(****************************************************************************************************<br>
© Syntegon Group.<br>
All rights reserved, also regarding any disposal, exploitation, reproduction, editing, distribution,<br>
as well as in the event of applications for industrial property rights.<br>
*****************************************************************************************************<br>
DESCRIPTION:<br>
Runtime-readable version of the Syn_Config library.<br>
*****************************************************************************************************<br>
VERSION         ¦ DATE       ¦ NAME      ¦ CHANGE<br>
Syn_Config 1.0.0 ¦ 2026-11-10 ¦ J.Willner ¦ Parameter sets of conveyors and Deltas (ADR 0017, protocol 1)<br>
Syn_Config 1.1.0 ¦ 2026-11-10 ¦ J.Willner ¦ Every other component type (#24)<br>
Syn_Config 2.0.0 ¦ 2026-11-11 ¦ J.Willner ¦ Gripper fingers in the robots' sets (protocol 2, #25)<br>
Syn_Config 2.0.1 ¦ 2026-11-12 ¦ J.Willner ¦ SynVisu as a placeholder: the application chooses its version<br>
Syn_Config 2.1.0 ¦ 2026-11-14 ¦ J.Willner ¦ Machine FB: recipe fields and machine commands (protocol 3, #43)<br>
Syn_Config 2.2.0 ¦ 2026-11-14 ¦ J.Willner ¦ Recipe fields: label, description, visibility condition (protocol 4, #49)<br>
Syn_Config 2.3.0 ¦ 2026-11-14 ¦ J.Willner ¦ One staging lifecycle; m_PassOn passes the pose on (Syn_Visu 10.0.0)<br>
Syn_Config 2.4.0 ¦ 2026-11-19 ¦ J.Willner ¦ Topology FB: nodes, roles and program links (protocol 5, #56)<br>
****************************************************************************************************)
FUNCTION _FC_GetVersionSynConfig : UINT
VAR_INPUT
	vi_n_VersionElement					: INT;	// [-] 1 = major, 2 = minor, 3 = revision
END_VAR

CASE vi_n_VersionElement OF
	1: _FC_GetVersionSynConfig := 2;
	2: _FC_GetVersionSynConfig := 4;
	3: _FC_GetVersionSynConfig := 0;
ELSE
	_FC_GetVersionSynConfig := 16#FFFF;
END_CASE

END_FUNCTION

(* stored: Version 1.1.0.1
   POU _FC_GetVersionSynConfig: Id {a7634710-508e-4100-adcb-bec076f572e5}, SpecialFunc None *)
